FUNCTION_BLOCK StandardMoverDetection IMPLEMENTS I_MoverDetectionAlgorithm
VAR
	iXtsTracks : ARRAY[0..TcIoXtsEnvironmentParameterList.MaxXtsTracksPerXpu] OF I_XtsTrack;
	iMoverArray : ARRAY[0..TcIoXtsEnvironmentParameterList.MaxXtsMoversPerXpu] OF I_XtsMover;
	iXPU : I_TcIoXtsProcessingUnit;
	XtsName : T_MaxString;
	MoverDetectionState : XtsMoverDetectionState;
	StartFlag : BOOL;
	ResetFlag : BOOL;
	_DetectedMoverCount: UDINT;
	MoverIdDetectionState: MoverIdDetectionStateEnum;
	MoverIdDetectionError: BOOL;
	MoverIdDetected: BOOL;
	_busy : BOOL;
	_done : BOOL;
	_error : BOOL;
END_VAR

{warning 'Add method implementation '}
METHOD Abort : HRESULT
END_METHOD

{warning 'Add property implementation'}
PROPERTY Busy : BOOL
GET
Busy := _busy;
END_GET
END_PROPERTY

METHOD Cycle : Base_Library.HRESULT
CASE MoverDetectionState OF
	XtsMoverDetectionState.WaitingForCommandStart:
		IF StartFlag THEN
			StartFlag := FALSE;
			_busy := TRUE;
			_done := FALSE;
			_error := FALSE;
			Base_Library.Tracing.Trace.Verbose(Source := XtsName, Message := 'Mover Detection Sequence Started');
			MoverDetectionState := XtsMoverDetectionState.SetATrackForDetection;
		END_IF
	XtsMoverDetectionState.SetATrackForDetection:
		Base_Library.Tracing.Trace.Verbose(Source := XtsName, Message := 'Track 1 set for detection');
		IXtsTracks[0].SetForDetection();
		MoverDetectionState := XtsMoverDetectionState.TriggeringRedetection;
	
	XtsMoverDetectionState.TriggeringRedetection:
		Base_Library.Tracing.Trace.Verbose(Source := XtsName, Message := 'Mover Redetection Started');
		IF iXPU.TriggerRedetection() THEN
			MoverDetectionState := XtsMoverDetectionState.WaitingForAllMoversValid;
		END_IF
		
	XtsMoverDetectionState.WaitingForAllMoversValid:
		IF iXPU.GetAreAllPositionsValid() THEN
			Base_Library.Tracing.Trace.Verbose(Source := XtsName, Message := 'All Movers Valid');
			MoverDetectionState := XtsMoverDetectionState.CheckingAllMoverFound;
		END_IF
	
	XtsMoverDetectionState.CheckingAllMoverFound:
		IF iXPU.GetExpectedMoverCount() = iXPU.GetDetectedMoverCount() THEN
			Base_Library.Tracing.Trace.Verbose(Source := XtsName, Message := 'Configured Movers = Detected Movers');
			_DetectedMoverCount := iXPU.GetDetectedMoverCount();
			MoverDetectionState := XtsMoverDetectionState.TriggeringMoverIdDetection;
		END_IF
		
	XtsMoverDetectionState.TriggeringMoverIdDetection:
		IF iXPU.GetMoverIdDetectionMode() = MoverIdDetectionMode.Standard OR_ELSE SUCCEEDED(TriggerMoverIDDetection()) THEN
			Base_Library.Tracing.Trace.Verbose(Source := XtsName, Message := 'Mover ID Detection Complete');
			MoverDetectionState := XtsMoverDetectionState.WaitingForCommandStart;
			_busy := FALSE;
			_done := TRUE;
		END_IF
		
	XtsMoverDetectionState.MoverDetectionFault:
		IF ResetFlag THEN
			ResetFlag := FALSE;
			_error := FALSE;
			MoverDetectionState := XtsMoverDetectionState.WaitingForCommandStart;
		END_IF
END_CASE
END_METHOD

PROPERTY DetectedMoverCount : UDINT
GET
DetectedMoverCount := _DetectedMoverCount;
END_GET
END_PROPERTY

{warning 'Add property implementation'}
PROPERTY Done : BOOL
GET
Done := _done;
END_GET
END_PROPERTY

{warning 'Add property implementation'}
PROPERTY Error : BOOL
GET
Error := _error;
END_GET
END_PROPERTY

PROPERTY Name : T_MAXSTRING
GET
END_GET
SET
XtsName := Name;
END_SET
END_PROPERTY

METHOD Reset : HRESULT
ResetFlag := TRUE;
END_METHOD

METHOD SetComponents : BOOL
VAR_INPUT
	XtsTracks : ARRAY[0..TcIoXtsEnvironmentParameterList.MaxXtsTracksPerXpu] OF I_XtsTrack;
	MoverArray : ARRAY[0..TcIoXtsEnvironmentParameterList.MaxXtsMoversPerXpu] OF I_XtsMover;
	XPU : I_TcIoXtsProcessingUnit;
END_VAR
iXtsTracks := XtsTracks;
iMoverArray := MoverArray;
iXPU := XPU;
END_METHOD

METHOD Start : HRESULT
StartFlag := TRUE;
END_METHOD

METHOD PRIVATE TriggerMoverIdDetection : HRESULT
VAR_INPUT
END_VAR
MoverIdDetectionError 	:= MoverIdDetectionState = MoverIdDetectionStateEnum.Error;
MoverIdDetected 	:= MoverIdDetectionState = MoverIdDetectionStateEnum.Valid;
MoverIdDetectionState	:= iXPU.GetMoverIdDetectionState();

IF iXPU.GetMoverIdDetectionMode() = MoverIdDetectionMode.Standard THEN
	TriggerMoverIDDetection := -1;
	RETURN;
END_IF
// 
IF MoverIdDetectionState = MoverIdDetectionStateEnum.Running THEN
	TriggerMoverIDDetection := -2;
	RETURN;
END_IF

iXPU.TriggerMoverIdDetection();
END_METHOD

END_FUNCTION_BLOCK

(* stored: Version 1.1.0.1
   POU StandardMoverDetection: Id {744247ae-04e1-4969-9309-29980f43d20b}, SpecialFunc None
   Method Abort: Id {26597c74-4029-447e-a786-072429fd8646}
   Property Busy: Id {7de3ebb0-a4b6-4ba8-a676-480469ee6c84}
   Get Get: Id {d94c0ad5-3b9d-4d0e-bb80-bdaaf09cfddb}
   Method Cycle: Id {ca7e54fe-ab1d-4501-9422-498d01d08e54}
   Property DetectedMoverCount: Id {8f21e2a7-94e9-4fac-bf40-130830a6435e}
   Get Get: Id {5b263380-d748-41dd-bfd1-9acc88eb9015}
   Property Done: Id {3c307923-0537-4387-97c5-91c7df94444f}
   Get Get: Id {61630dd0-000e-4a6d-b174-fb82efe87251}
   Property Error: Id {49b9de1e-4304-4b08-b048-a12a8d110617}
   Get Get: Id {99b1ff45-eeef-414e-b891-4cb8cddc003e}
   Property Name: Id {d6ec0b86-8dd6-4548-b7b5-ce4cb41bc7bc}
   Get Get: Id {eeb06967-34c8-4544-b485-ab92c5ed582c}
   Set Set: Id {9752c199-4b0a-4393-aefb-b87162e2ed87}
   Method Reset: Id {4debf444-f915-47ef-8621-fa026afbedd9}
   Method SetComponents: Id {85ce5b9a-63bb-4bb2-bedb-42a81ea16fe0}
   Method Start: Id {507dae7d-fc01-4c32-8358-312d0dae6a9b}
   Method TriggerMoverIdDetection: Id {49e4cae6-2a7e-45cb-ba80-e12b965b943f} *)
